// TIA Portal V21 export
FUNCTION_BLOCK "GraphQualification"   // FB, GRAPH
// stored: AutoNumber true
   VAR_INPUT
      ACK_EF : Bool;
   END_VAR
BEGIN
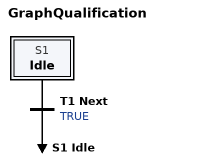
   // sequencer 1
   INITIAL_STEP Idle:   // S1
   END_STEP
   TRANSITION Next FROM Idle TO Idle   // T1, jump
      := TRUE;
   END_TRANSITION
END_FUNCTION_BLOCK
